Fanuc KAREL source: KA00080.KL

PROGRAM KA00080
%NOLOCKGROUP
VAR
  SRC: XYZWPREXT
  DST: JOINTPOS
BEGIN
  SRC.X = 1.0
  DST = SRC
END KA00080
